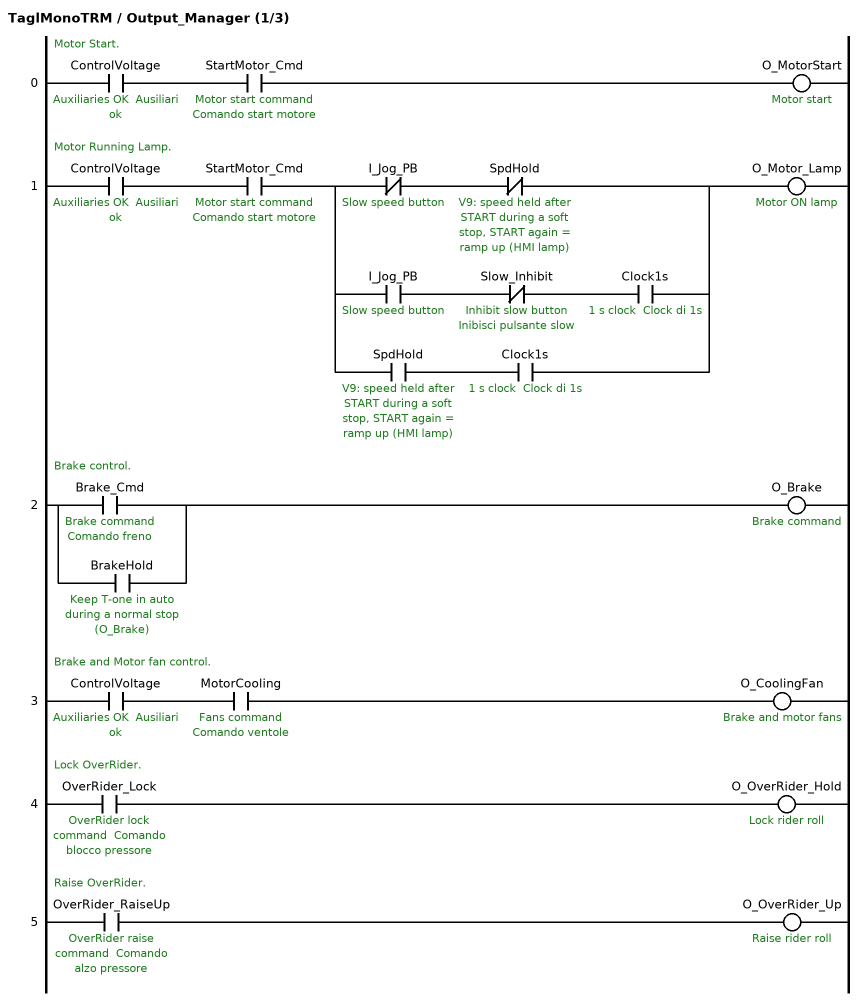
(* [picture p24: TaglMonoTRM / Output_Manager, rungs 0-5] *)
(* Rung 0: Motor Start. *)
O_MotorStart := ControlVoltage AND StartMotor_Cmd;
(* Rung 1: Motor Running Lamp. *)
O_Motor_Lamp := ControlVoltage AND StartMotor_Cmd AND ((NOT I_Jog_PB AND NOT SpdHold) OR (I_Jog_PB AND NOT Slow_Inhibit AND Clock1s) OR (SpdHold AND Clock1s));
(* Rung 2: Brake control. *)
O_Brake := Brake_Cmd OR BrakeHold;
(* Rung 3: Brake and Motor fan control. *)
O_CoolingFan := ControlVoltage AND MotorCooling;
(* Rung 4: Lock OverRider. *)
O_OverRider_Hold := OverRider_Lock;
(* Rung 5: Raise OverRider. *)
O_OverRider_Up := OverRider_RaiseUp;

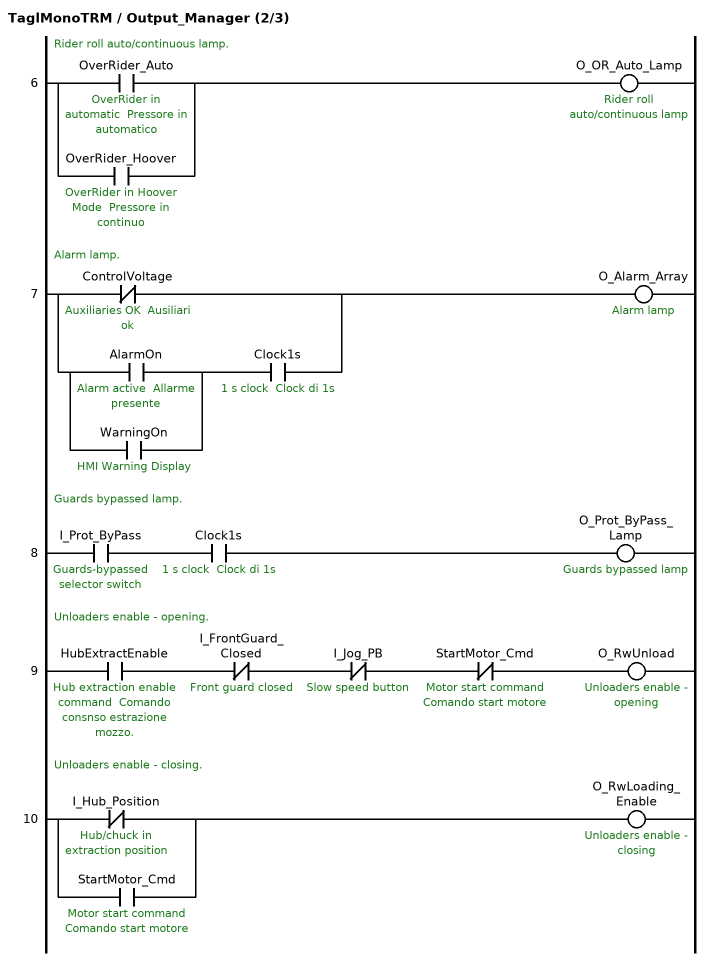
(* Rung 6: Rider roll auto/continuous lamp. *)
O_OR_Auto_Lamp := OverRider_Auto OR OverRider_Hoover;
(* Rung 7: Alarm lamp. *)
O_Alarm_Array := NOT ControlVoltage OR ((AlarmOn OR WarningOn) AND Clock1s);
(* Rung 8: Guards bypassed lamp. *)
O_Prot_ByPass_Lamp := I_Prot_ByPass AND Clock1s;
(* Rung 9: Unloaders enable - opening. *)
O_RwUnload := HubExtractEnable AND NOT I_FrontGuard_Closed AND NOT I_Jog_PB AND NOT StartMotor_Cmd;
(* Rung 10: Unloaders enable - closing. *)
O_RwLoading_Enable := NOT I_Hub_Position OR StartMotor_Cmd;

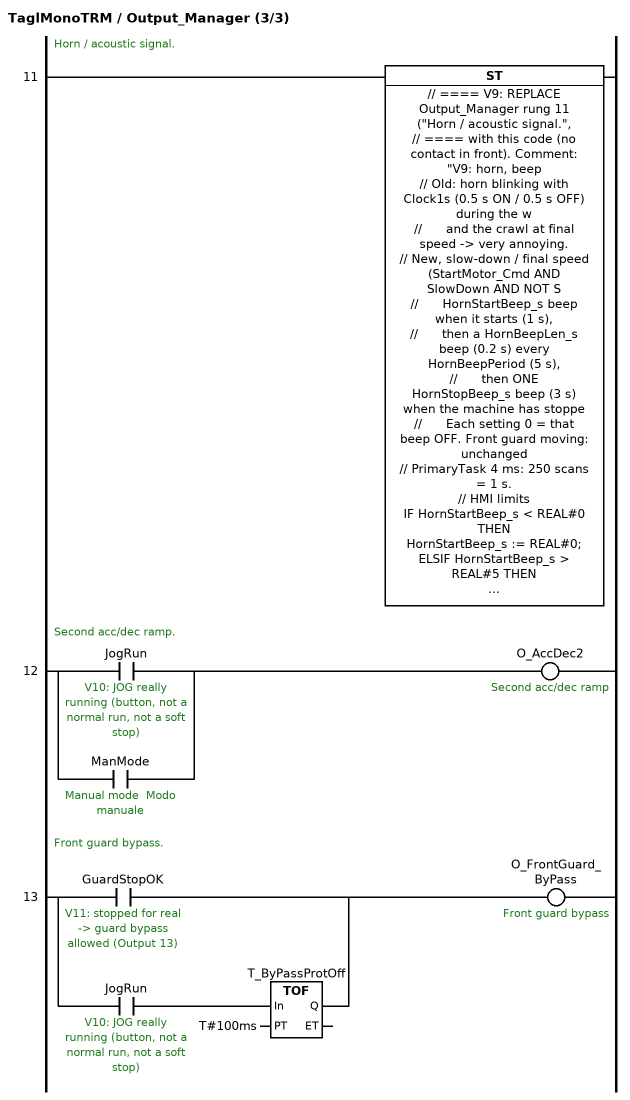
(* Rung 11: Horn / acoustic signal. *)
// ==== V9: REPLACE Output_Manager rung 11 ("Horn / acoustic signal.", ladder) by ONE ST rung
// ==== with this code (no contact in front). Comment: "V9: horn, beeps set on the HMI".
// Old: horn blinking with Clock1s (0.5 s ON / 0.5 s OFF) during the whole slow-down
//      and the crawl at final speed -> very annoying.
// New, slow-down / final speed (StartMotor_Cmd AND SlowDown AND NOT Stop):
//      HornStartBeep_s beep when it starts (1 s),
//      then a HornBeepLen_s beep (0.2 s) every HornBeepPeriod (5 s),
//      then ONE HornStopBeep_s beep (3 s) when the machine has stopped (< 2 m/min).
//      Each setting 0 = that beep OFF. Front guard moving: unchanged (Clock1s blinking).
// PrimaryTask 4 ms: 250 scans = 1 s.

// HMI limits

IF HornStartBeep_s < REAL#0 THEN
    HornStartBeep_s := REAL#0;
ELSIF HornStartBeep_s > REAL#5 THEN
    HornStartBeep_s := REAL#5;
END_IF;

IF HornBeepLen_s < REAL#0 THEN
    HornBeepLen_s := REAL#0;
ELSIF HornBeepLen_s > REAL#2 THEN
    HornBeepLen_s := REAL#2;
END_IF;

IF HornBeepPeriod < REAL#0 THEN
    HornBeepPeriod := REAL#0;
ELSIF (HornBeepPeriod > REAL#0) AND (HornBeepPeriod < HornBeepLen_s + REAL#0.5) THEN
    HornBeepPeriod := HornBeepLen_s + REAL#0.5;     // always a pause between beeps
ELSIF HornBeepPeriod > REAL#30 THEN
    HornBeepPeriod := REAL#30;
END_IF;

IF HornStopBeep_s < REAL#0 THEN
    HornStopBeep_s := REAL#0;
ELSIF HornStopBeep_s > REAL#10 THEN
    HornStopBeep_s := REAL#10;
END_IF;

HornStartScans := REAL_TO_INT(HornStartBeep_s * REAL#250);
HornLenScans   := REAL_TO_INT(HornBeepLen_s * REAL#250);
HornPer        := REAL_TO_INT(HornBeepPeriod * REAL#250);

// Slow-down / final speed beeps

HornRun := StartMotor_Cmd AND SlowDown AND NOT Stop;

IF HornRun THEN
    IF NOT HornRunMem THEN
        HornTicks := 0;                             // slow-down starts
    END_IF;
	
    IF HornTicks < 30000 THEN
        HornTicks := HornTicks + 1;
    END_IF;
	
    IF HornTicks <= HornStartScans THEN
        HornSlowBeep := TRUE;                       // start beep
        HornCnt := 0;
    ELSIF (HornPer > 0) AND (HornLenScans > 0) THEN
        HornCnt := HornCnt + 1;
        IF HornCnt >= HornPer THEN
            HornCnt := 0;
        END_IF;
		
        HornSlowBeep := (HornCnt >= HornPer - HornLenScans);   // beep at the end of each period
    ELSE
        HornSlowBeep := FALSE;                      // periodic beeps OFF
    END_IF;
ELSE
    HornTicks := 0;
    HornCnt := 0;
    HornSlowBeep := FALSE;
END_IF;

// End of a slow-down by a stop (auto stop, STOP button): one beep at standstill
// (Stop is set in Motor_Manager before StartMotor_Cmd drops on the next scan)

IF HornRunMem AND NOT HornRun AND (Stop OR NOT StartMotor_Cmd) THEN
    HornStopPend := TRUE;
END_IF;

IF StartMotor_Cmd AND NOT HornStartMem THEN
    HornStopPend := FALSE;                          // restarted: no stop beep
    HornStopTicks := 0;
END_IF;

HornStartMem := StartMotor_Cmd;

IF HornStopPend AND (Velocity_M_min < REAL#2) THEN
    HornStopPend := FALSE;
    HornStopTicks := REAL_TO_INT(HornStopBeep_s * REAL#250);
END_IF;

IF HornStopTicks > 0 THEN
    HornStopTicks := HornStopTicks - 1;
END_IF;

HornRunMem := HornRun;

// HMI test button: horn while pressed (machine stopped only)

O_AcousticSignal := (NOT I_FrontGuard_Closed AND NOT I_FrontGuard_Open AND Clock1s)
                    OR HornSlowBeep OR (HornStopTicks > 0)
                    OR (HornTest AND NOT StartMotor_Cmd);
(* Rung 12: Second acc/dec ramp. *)
O_AccDec2 := JogRun OR ManMode;
(* Rung 13: Front guard bypass. *)
T_ByPassProtOff(In := JogRun, PT := T#100ms);
O_FrontGuard_ByPass := GuardStopOK OR T_ByPassProtOff.Q;

(* Section AutoStop_Control: ladder, written here as Structured Text *)

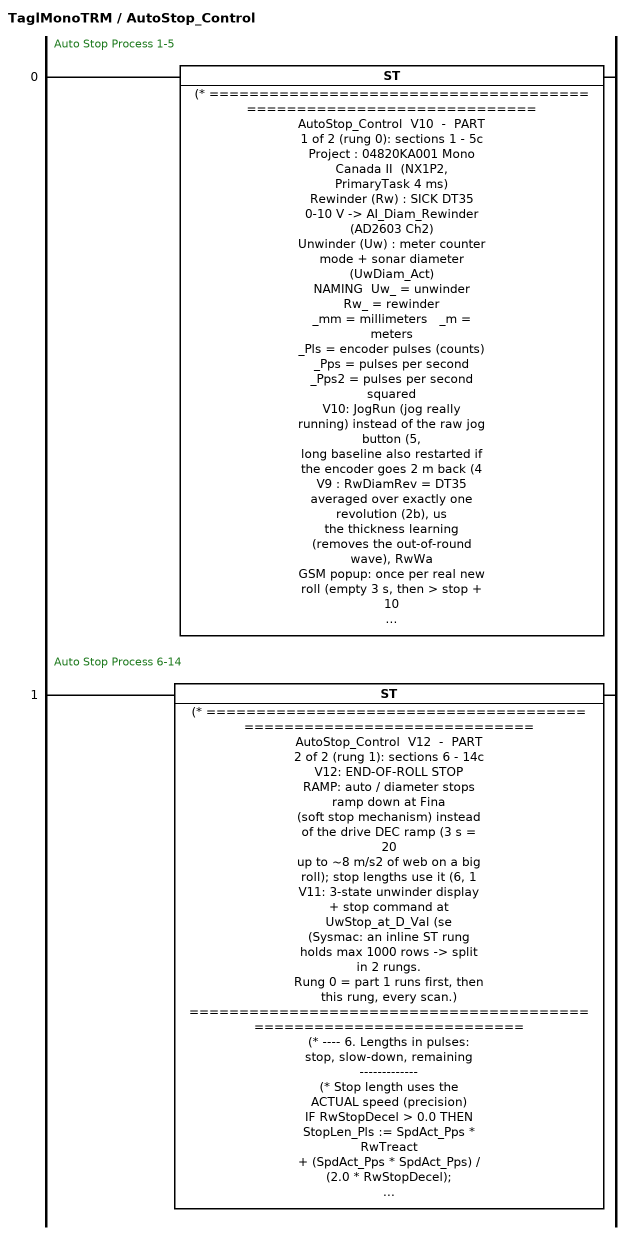
(* Rung 0: Auto Stop Process 1-5 *)
(* ==========================================================================
   AutoStop_Control  V10  -  PART 1 of 2 (rung 0): sections 1 - 5c
   Project : 04820KA001 Mono Canada II  (NX1P2, PrimaryTask 4 ms)
   Rewinder (Rw) : SICK DT35 0-10 V -> AI_Diam_Rewinder (AD2603 Ch2)
   Unwinder (Uw) : meter counter mode + sonar diameter (UwDiam_Act)

   NAMING  Uw_ = unwinder   Rw_ = rewinder
           _mm = millimeters   _m = meters
           _Pls = encoder pulses (counts)   _Pps = pulses per second
           _Pps2 = pulses per second squared

   V10: JogRun (jog really running) instead of the raw jog button (5, 5b);
          long baseline also restarted if the encoder goes 2 m back (4b).
   V9 : RwDiamRev = DT35 averaged over exactly one revolution (2b), used by
          the thickness learning (removes the out-of-round wave), RwWave_mm.
        GSM popup: once per real new roll (empty 3 s, then > stop + 100 mm
          for 3 s); NEW PAPER closes it (section 10).
        paper thickness: long-baseline learning (D^2 growth / length) from the
          start point, LOCKED at RwLockDiam (300 mm): no more change, no
          paper-change detection, until NEW PAPER / GSM popup YES (4b).
   V8 : = V7 + V7c unwinder DIAMETER slow-down follows the speed (6c),
          V7e ManMode slow-down model as before V7 (section 6),
          V7f S-curve extra length in the slow-down (section 6)
   V7 : FEED-FORWARD speed loop (Motor_Manager rung B): reference = set speed
        x RwRatioD / diameter along a ramp in real web mm/s2 (DecelWeb /
        AccelWeb), RwRatioD adapted slowly -> no hunting on big rolls.
        Section 6: slow-down length = one ramp at DecelWeb (FFEnable), else
        web coarse ramp + trim tail; learning only as fallback.
   v6y: rewinder AUTO stop (RwStopEnable) limits the work speed to
        RwAutoMaxSpd (500 m/min), taken over at standstill only; section 6
        uses the limited speed.
   v6x: new parent roll on the unwinder -> GsmAsk (HMI popup "did you change
        the paper?"); GsmAskYes forgets the learned thickness.
   v6w: paper thickness window is LENGTH-based instead of 10 s, modulated by
        the diameter (RwWinGrow_mm 2.5 mm of growth, 4 m .. RwWinLen_m 30 m):
        same accuracy at every speed and roll size; stopped window = dropped.
        ALARM RESET also clears LearnFailCnt / StopFailCnt (alarm 16).
   v6v: BrakeHold released on the SIGNED web speed (Velocity_M_min < 5),
        so a web pulled back after the stop releases the T-one at once.
   v6u: stop learning: a stop shorter than the reaction distance or faster
        than RwDecelMax_mm is ignored (not a fault). Only a too slow stop
        (< RwDecelMin_mm) counts toward alarm 16.
   v6t: rewinder slow-down fallback while the paper thickness is not
        learned: RwSlowReq at RwTargetDiam - RwSlowFallbackMm (30 mm).
   v6s: paper change: a learning window more than RwMatChangePct (25 %) away
        from RwMat_K is ignored once, taken directly the 2nd time in a row
        (automatic). RwMatReset (HMI "NEW PAPER") forgets RwMat_K.
   v6p: section 5c: RwLearnReset clears RwStopDecelK, RwStopDecel and
        RwSlowDecelK (the v6f seed that refilled RwStopDecelK is removed).
   v6l: previous value saved before every TEACH CORE (RwAxisDist_Prev,
          UwCoreDist_Prev, Retain) + UNDO buttons (RwTeachUndo,
          UwTeachUndo): swap current <-> previous. State 4 = RESTORED.
   v6k: unwinder TEACH CORE (Core_Measure) works like the rewinder one:
          same checks, 2 s stable with sonar AVERAGE, status UwTeachState.
          Replaces General rung 15 (one immediate sonar reading).
   v6j: TEACH CORE (section 14): HMI button RwTeachCore, empty core on the
          rewinder, machine stopped -> after 2 s stable:
          RwAxisDist := RwDist + RwCoreDiameter / 2. Status in RwTeachState.
   v6i: auto: pots scaled to WorkSpd_Max / FinalSpd_Max (Motor_Manager rung 6,
          Pot1_Mem / Pot2_Mem). ManMode keeps the raw pots (percent),
          so section 6 uses the raw pots in ManMode.
   v6h: BrakeHold keeps O_Brake (T-one "reel brake automatic") ON during a
          normal stop until the web is almost stopped (< 5 m/min, max 15 s).
          Before: T-one switched to "stop" with the run command, while the
          rewinder was decelerating hard -> unwinder overran, web on the
          floor (field 10/20/2026). Used in Output_Manager rung 2.
   v6g: slow-down AND stop decel proportional to the rewinder diameter.
          The ATV930 ramp is in Hz/s (motor = rewind shaft), so the web
          decel [mm/s2] = shaft decel x radius. Field data 10/20/2026:
          24 mm/s2 at 120 mm -> 90 mm/s2 at 600 mm.
          Learned: RwSlowDecelK, RwStopDecelK [mm/s2 per mm of diameter].
          Live:    RwSlowDecelLrn [mm/s2], RwStopDecel [pulses/s2] = K x DecelDiam.
   v6f: learn the REAL slow-down deceleration (section 5b) -> RwSlowDecelLrn
          (mm/s2). The ATV930 stretches its ramp with a heavy roll (no
          braking resistor), so the PLC ramp (DecelCoarse) was too
          optimistic: the stop came before final speed was reached.
          Priority in section 6: RwSlowDecel (manual) > RwSlowDecelLrn
          (learned) > DecelCoarse/DecelTrim model.
   v6e: GSM_Learned_OK (replaces global RwLearnFault): TRUE only when
          RwMat_K is learned, RwStopDecel is learned (if RwLearnStop) and
          there is no learning fault. Alarm 16 uses GSM_LearnFault.
   v6d: exact 100 ms tick (25 x 4 ms scan counter, the self-resetting
          TON ran ~104-108 ms -> speed ~4-8 % too high)
        standstill = <= 2 counts / 100 ms (encoder jitter)
        stop learning skipped after jog / manual / slow-button runs and
          when the auxiliaries drop (E-stop): RunWasJog, StopLearnValid
        work / final speed from the potentiometers in BOTH modes
          (Speed_Display / LowSpd_Display are not m/min in ManMode)
        slow-down length includes the DecelTrim tail inside the
          SpdDelta_Percent band (Motor_Manager rungs 14/15)
   v6c: learning supervision -> RwLearnFault (alarm 16), learned paper
          thickness RwThick_mm, plausibility limits for K and stop decel
   v6b: RwMaxSlowAtDiam display + RwMaxSlowFallback (slow-down warning
          while RwMat_K is not learned yet)
   v6 : consistent internal names, units in names.
        Globals renamed: RwRemain_m, RwStopLen_m, RwSlowLen_m,
                         RwSlowMargin_m, UwSlowMargin_m
   v5 : max diameter protection (always active), sensor plausibility,
        12SA5 master (section 9), alarms in section Alarms (ladder)
   v4b: AUTO interlock + single HMI display (SlowAtDisp / SlowAtMode)
   ========================================================================== *)

(* ---- 1. 100 ms tick, mm per encoder pulse ------------------------------ *)
(* v6d: 25 scans x 4 ms PrimaryTask = exactly 100 ms.                       *)
(*      Change 25 if the PrimaryTask period is changed.                    *)

TickCnt := TickCnt + 1;

IF TickCnt >= 25 THEN
    TickCnt := 0;
    Tick := TRUE;
ELSE
    Tick := FALSE;
END_IF;

IF (Encoder_Pulse > 0) AND (EncoderWheel_Circumf > 0.0) THEN
    MmPerPulse := EncoderWheel_Circumf / (INT_TO_REAL(Encoder_Pulse) * 4.0);
ELSE
    MmPerPulse := 0.0;
END_IF;

(* ---- 2. Rewinder DT35 -> filtered distance -> diameter ----------------- *)

RwDistRaw_mm := RwDist0V + (INT_TO_REAL(AI_Diam_Rewinder) / 4000.0)
                * (RwDist10V - RwDist0V);

IF Tick THEN
    IF NOT RwFiltInit THEN
        RwDist := RwDistRaw_mm;
        RwFiltInit := TRUE;
    ELSE
        RwDist := RwDist + RwFilter_K * (RwDistRaw_mm - RwDist);
    END_IF;
END_IF;

RwSensFault := (AI_Diam_Rewinder < RwRawMin) OR (AI_Diam_Rewinder > RwRawMax)
               OR (RwDist > RwAxisDist);

RwDiam := 2.0 * (RwAxisDist - RwDist);

IF RwDiam < 0.0 THEN
    RwDiam := 0.0;
END_IF;

(* ---- 2b. V9: diameter averaged over exactly ONE revolution -------------- *)
(* The out-of-round roll gives a wave at the rotation frequency (seen in   *)
(* the 10/29 traces: 2.4 Hz at 444 m/min / 973 mm). Averaging the raw     *)
(* DT35 distance over exactly one revolution cancels it (and all its      *)
(* harmonics), whatever the phase -> no shaft position sensor needed:     *)
(* one revolution = PI x D of web on the encoder. Each scan is weighted   *)
(* by its encoder pulses = by roll ANGLE, so ramps and standstill do not  *)
(* bias it (stopped: nothing added). Used only by the thickness learning. *)
(* RwWave_mm = peak-peak diameter wave in the last revolution (HMI).      *)

RevDP := ABS(Encoder_Pos - RevPrevPos);
RevPrevPos := Encoder_Pos;

IF RwSensFault OR (MmPerPulse <= 0.0) OR (RwDiam < 50.0) OR (RevDP > 100000) THEN
    RevW := 0.0;
    RevSum := 0.0;
    RwDiamRevOk := RwDiamRevOk AND NOT RwSensFault;
ELSIF RevDP > 0 THEN
	
    IF RevW <= 0.0 THEN
        RevMin := RwDistRaw_mm;
        RevMax := RwDistRaw_mm;
    END_IF;
	
    RevSum := RevSum + RwDistRaw_mm * DINT_TO_REAL(RevDP);
    RevW := RevW + DINT_TO_REAL(RevDP);
	
    IF RwDistRaw_mm < RevMin THEN
        RevMin := RwDistRaw_mm;
    END_IF;
	
    IF RwDistRaw_mm > RevMax THEN
        RevMax := RwDistRaw_mm;
    END_IF;
	
    IF RevW >= 3.14159 * RwDiam / MmPerPulse THEN
        RwDiamRev := 2.0 * (RwAxisDist - RevSum / RevW);
        RwWave_mm := 2.0 * (RevMax - RevMin);
        RwDiamRevOk := TRUE;
        RevW := 0.0;
        RevSum := 0.0;
    END_IF;
END_IF;

(* v6g: diameter used by the decel model (last valid on sensor fault)      *)

IF NOT RwSensFault THEN
    DecelDiam := RwDiam;
ELSE
    DecelDiam := RwLastValidDiam;
END_IF;

IF DecelDiam < 100.0 THEN
    DecelDiam := 100.0;                             (* core *)
END_IF;

(* ---- 3. Actual speed from encoder, 100 ms window ----------------------- *)

IF Tick THEN
	
    IF NOT SpdInit THEN
        EncPrev := Encoder_Pos;
        SpdInit := TRUE;
    END_IF;
	
    SpdAct_Pps := DINT_TO_REAL(ABS(Encoder_Pos - EncPrev)) * 10.0;
    EncPrev := Encoder_Pos;
END_IF;

RwSpeed := SpdAct_Pps * MmPerPulse * 0.06;          (* m/min *)

(* ---- 4a. v6s: NEW PAPER button: forget the learned thickness ----------- *)
(* RwMat_K = 0 -> the first valid 10 s window sets it directly.            *)
(* HMI momentary button: must be HELD 3 s, then the reset is done once and *)
(* the PLC clears the bit (HMI lamp goes off = done).                      *)

T_MatReset(In := RwMatReset, PT := T#3s);

IF T_MatReset.Q THEN
    RwMat_K := 0.0;
    LearnFailCnt := 0;
    MatChangeCnt := 0;
    RwMatLocked := FALSE;                           (* V9 *)
    LongActive := FALSE;
    GsmAsk := FALSE;                                (* V9: NEW PAPER answers the popup *)
    GsmArmed := FALSE;
    RwMatReset := FALSE;
END_IF;

(* ---- 4b. V9: long-baseline thickness learning + LOCK ------------------- *)
(* From the start point (first run after NEW PAPER / GSM YES / power-on    *)
(* while not locked): K = (D^2 - D0^2) / (2 x pulses). The waving of the   *)
(* roll (+/-0.4 mm) only matters at the two ends, so the error falls with  *)
(* the growth (50 mm growth: ~1 %). After 20 mm growth it replaces the     *)
(* 30 m windows. At RwLockDiam (and >= RwLockMinGrow_mm growth) the value *)
(* is LOCKED (Retain): windows and paper-change detection stop.            *)
(* RwLockDiam = 0 -> never locked (windows + long baseline as learning).   *)

IF Tick AND NOT RwMatLocked THEN
	
    IF LongActive AND (RwDiamRev < LongStartD - 30.0) AND RwDiamRevOk THEN
        LongActive := FALSE;                        (* new core: restart *)
    END_IF;
	
    IF Encoder_Reset OR (Encoder_Pos < LongStartPos - 20000) THEN
        LongActive := FALSE;                        (* metre counter reset / 2 m back *)
    END_IF;
	
    IF NOT LongActive AND O_MotorStart AND RwDiamRevOk
       AND (RwDiamRev > 0.0) THEN
        LongStartPos := Encoder_Pos;
        LongStartD := RwDiamRev;
        LongActive := TRUE;
    END_IF;
	
    LongValid := FALSE;
	
    IF LongActive AND RwDiamRevOk AND (MmPerPulse > 0.0) THEN
        LongGrow_mm := RwDiamRev - LongStartD;
        LongPls := DINT_TO_REAL(ABS(Encoder_Pos - LongStartPos));
		
        IF (LongGrow_mm >= 20.0) AND (LongPls > 0.0) THEN
            LongK := (RwDiamRev * RwDiamRev - LongStartD * LongStartD) / (2.0 * LongPls);
            LongThick_mm := LongK * 3.14159 / (2.0 * MmPerPulse);
			
            IF (LongThick_mm >= RwThickMin_mm) AND (LongThick_mm <= RwThickMax_mm) THEN
                LongValid := TRUE;
                RwMat_K := LongK;
                MatChangeCnt := 0;
                LearnFailCnt := 0;
				
                IF (RwLockDiam > 0.0) AND (RwDiamRev >= RwLockDiam)
                   AND (LongGrow_mm >= RwLockMinGrow_mm) THEN
                    RwMatLocked := TRUE;            (* solid from now on *)
                    LongActive := FALSE;
                END_IF;
            END_IF;
        END_IF;
    END_IF;
END_IF;

IF RwMatLocked THEN
    LongValid := FALSE;
    LearnFailCnt := 0;                              (* no thickness alarm *)
END_IF;

(* ---- 4. Learn material factor  K = dDiam/dPulse * Diam ----------------- *)

IF Tick THEN
    LearnWinTicks := LearnWinTicks + 1;
	
    IF NOT LearnInit THEN
        LearnWinStartPos := Encoder_Pos;  LearnWinStartDiam := RwDiamRev;  (* V9 *)
        LearnWinTicks := 0;
        LearnWinRunning := O_MotorStart;
        LearnInit := TRUE;
    ELSE
        LearnWinRunning := LearnWinRunning AND O_MotorStart;
        (* v6w: LENGTH-based window, modulated by the diameter: closes    *)
        (* when the roll should have grown RwWinGrow_mm (2.5 mm), so the  *)
        (* accuracy vs DT35 noise is the same at every speed and size.    *)
        (* Pulses = growth x diameter / K (K = learned RwMat_K).          *)
        (* Limits: min 4 m, max RwWinLen_m (30 m). K not learned: max.    *)
        (* Motor stopped during the window -> window dropped (no fault).  *)
		
        IF MmPerPulse > 0.0 THEN
            IF (RwMat_K > 0.0) AND (RwWinGrow_mm > 0.0) THEN
                LearnWinLen_Pls := RwWinGrow_mm * MAX(RwDiam, REAL#100.0) / RwMat_K;
            ELSE
                LearnWinLen_Pls := RwWinLen_m * 1000.0 / MmPerPulse;
            END_IF;
			
            IF LearnWinLen_Pls < 4000.0 / MmPerPulse THEN
                LearnWinLen_Pls := 4000.0 / MmPerPulse;              (* 4 m *)
            END_IF;
			
            IF (RwWinLen_m > 0.0)
               AND (LearnWinLen_Pls > RwWinLen_m * 1000.0 / MmPerPulse) THEN
                LearnWinLen_Pls := RwWinLen_m * 1000.0 / MmPerPulse;
            END_IF;
        ELSE
            LearnWinLen_Pls := 300000.0;
        END_IF;
		
        IF (DINT_TO_REAL(ABS(Encoder_Pos - LearnWinStartPos)) >= LearnWinLen_Pls)
           OR NOT LearnWinRunning THEN
            LearnWin_Pls := ABS(Encoder_Pos - LearnWinStartPos);
            LearnWinDiamDelta := RwDiamRev - LearnWinStartDiam;  (* V9 *)
            (* A window SHOULD learn: ran all the time, enough length,  *)
            (* DT35 OK. Then it must give a plausible paper thickness. *)
			
            IF LearnWinRunning AND (LearnWin_Pls >= RwMinPulses)
               AND NOT RwSensFault
               AND NOT RwMatLocked AND NOT LongValid      (* V9 *)
               AND RwDiamRevOk AND (LearnWinStartDiam > 0.0) THEN
                LearnWinOk := FALSE;
				
                IF (LearnWinDiamDelta > 0.0) AND (MmPerPulse > 0.0) THEN
                    MatK_Window := (LearnWinDiamDelta / DINT_TO_REAL(LearnWin_Pls))
                                   * ((RwDiamRev + LearnWinStartDiam) / 2.0);
                    (* K = 2 * thickness * mm-per-pulse / PI          *)
                    ThickWin_mm := MatK_Window * 3.14159 / (2.0 * MmPerPulse);
					
                    IF (ThickWin_mm >= RwThickMin_mm)
                       AND (ThickWin_mm <= RwThickMax_mm) THEN
                        LearnWinOk := TRUE;
						
                        IF RwMat_K <= 0.0 THEN
                            RwMat_K := MatK_Window;
                            MatChangeCnt := 0;
                        ELSIF (RwMatChangePct > 0.0)
                              AND (ABS(MatK_Window - RwMat_K)
                                   > RwMat_K * RwMatChangePct / 100.0) THEN
                            (* v6s: far from the learned value: 1 window = ignored *)
                            (* (outlier), 2 in a row = paper changed -> take it.  *)
                            MatChangeCnt := MatChangeCnt + 1;
							
                            IF MatChangeCnt >= 2 THEN
                                RwMat_K := MatK_Window;
                                MatChangeCnt := 0;
                            END_IF;
                        ELSE
                            MatChangeCnt := 0;
                            RwMat_K := RwMat_K + RwLearn_K * (MatK_Window - RwMat_K);
                        END_IF;
                    END_IF;
                END_IF;
				
                IF LearnWinOk THEN
                    LearnFailCnt := 0;
                ELSIF LearnFailCnt < 1000 THEN
                    LearnFailCnt := LearnFailCnt + 1;  (* no growth / implausible *)
                END_IF;
            END_IF;
            LearnWinStartPos := Encoder_Pos;  LearnWinStartDiam := RwDiamRev;  (* V9 *)
            LearnWinTicks := 0;
            LearnWinRunning := O_MotorStart;
        END_IF;
    END_IF;
END_IF;

(* ---- 5. Learn real stop deceleration on every stop --------------------- *)
(* v6d: a run with jog / manual / slow button uses the 2nd ramp (O_AccDec2) *)
(*      -> its stop must not be learned. Latched for the whole run because  *)
(*      the jog button is already released on the stop edge.                  *)

IF O_MotorStart AND NOT MotorRunMem THEN            (* start edge *)
    RunWasJog := FALSE;
END_IF;

IF O_MotorStart AND (ManMode OR JogRun) THEN
    RunWasJog := TRUE;
END_IF;

IF MotorRunMem AND NOT O_MotorStart THEN            (* stop command edge *)
    StopMeasActive := TRUE;
    StopStartPos := Encoder_Pos;
    StopStartSpd_Pps := SpdAct_Pps;
    StopStartDiam := DecelDiam;
    StandstillTicks := 0;
    (* STOP button and automatic stop take the same path (drive DI1 and    *)
    (* O_Brake -> T-one drop together, electrical plan sheets 1/9/15),     *)
    (* so both are learned.                                                *)
    StopLearnValid := ControlVoltage AND NOT RunWasJog AND NOT ManMode;
END_IF;

MotorRunMem := O_MotorStart;

IF O_MotorStart THEN
    StopMeasActive := FALSE;                        (* restarted: abort *)
ELSIF StopMeasActive AND Tick THEN
	
    IF NOT ControlVoltage THEN
        StopLearnValid := FALSE;                    (* E-stop during the stop *)
    END_IF;
	
    IF SpdAct_Pps <= 20.0 THEN                      (* <= 2 counts / 100 ms *)
        StandstillTicks := StandstillTicks + 1;
    ELSE
        StandstillTicks := 0;
    END_IF;
	
    IF StandstillTicks >= 3 THEN                    (* standstill 300 ms *)
        StopMeasActive := FALSE;
        StopMeas_Pls := DINT_TO_REAL(ABS(Encoder_Pos - StopStartPos));
		
        IF RwLearnStop AND StopLearnValid
           AND (StopStartSpd_Pps * MmPerPulse * 0.06 >= RwMinLearnSpd) THEN
            (* This stop SHOULD learn: result must be plausible       *)
            (* v6u: a stop shorter than the reaction distance, or     *)
            (* faster than RwDecelMax_mm, is NOT a fault: the web      *)
            (* stopped within a few mm, nothing to learn (trace        *)
            (* 10/28/2026: 23 m/min -> stopped in 102 pulses = 10 mm). *)
            (* Only a too SLOW stop (< RwDecelMin_mm) counts as fail.  *)
            StopLearnOk := FALSE;
			
            IF StopMeas_Pls > StopStartSpd_Pps * RwTreact THEN
                StopDecelMeas := (StopStartSpd_Pps * StopStartSpd_Pps)
                                 / (2.0 * (StopMeas_Pls - StopStartSpd_Pps * RwTreact));
                StopDecelMeas_mm := StopDecelMeas * MmPerPulse;  (* mm/s2 *)
				
                IF (StopDecelMeas_mm >= RwDecelMin_mm)
                   AND (StopDecelMeas_mm <= RwDecelMax_mm) THEN
                    StopLearnOk := TRUE;
                    (* v6g: learn per mm of diameter *)
                    DecelK_Meas := StopDecelMeas_mm / ((StopStartDiam + DecelDiam) / 2.0);
					
                    IF RwStopDecelK <= 0.0 THEN
                        RwStopDecelK := DecelK_Meas;
                    ELSE
                        RwStopDecelK := RwStopDecelK + 0.3 * (DecelK_Meas - RwStopDecelK);
                    END_IF;
					
                    StopFailCnt := 0;
                ELSIF StopDecelMeas_mm < RwDecelMin_mm THEN
					
                    IF StopFailCnt < 1000 THEN
                        StopFailCnt := StopFailCnt + 1;    (* stop too long *)
                    END_IF;
                END_IF;                                    (* too fast: ignored *)
            END_IF;                                        (* too short: ignored *)
        END_IF;
    END_IF;
END_IF;

(* ---- 5b. v6f: learn real slow-down deceleration ----------------------- *)
(* From the SlowDown edge (at speed) until final speed is reached, or     *)
(* until the stop comes first. a = (v0^2 - v1^2) / (2 * distance).         *)
(* Not learned in jog / manual / slow button (2nd ramp).                   *)

IF SlowDown AND NOT SlowMem AND O_MotorStart
   AND NOT ManMode AND NOT JogRun
   AND (SpdAct_Pps > SpdFinal_Pps + SpdBand_Pps) THEN
    SlowMeasActive := TRUE;
    SlowStartPos := Encoder_Pos;
    SlowStartSpd_Pps := SpdAct_Pps;
    SlowStartDiam := DecelDiam;
END_IF;
SlowMem := SlowDown;

IF SlowMeasActive THEN
	
    IF NOT SlowDown OR ManMode OR JogRun THEN
        SlowMeasActive := FALSE;                    (* aborted *)
    ELSIF Tick AND ((SpdAct_Pps <= SpdFinal_Pps + 0.25 * SpdBand_Pps)
                    OR NOT O_MotorStart) THEN       (* final reached or stopped *)
        SlowMeasActive := FALSE;
        SlowMeas_Pls := DINT_TO_REAL(ABS(Encoder_Pos - SlowStartPos));
		
        IF (SlowMeas_Pls > 0.0) AND (MmPerPulse > 0.0)
           AND ((SlowStartSpd_Pps - SpdAct_Pps) * MmPerPulse * 0.06 >= 10.0) THEN
            SlowDecelMeas_mm := (SlowStartSpd_Pps * SlowStartSpd_Pps
                                 - SpdAct_Pps * SpdAct_Pps)
                                / (2.0 * SlowMeas_Pls) * MmPerPulse;  (* mm/s2 *)
								
            IF (SlowDecelMeas_mm >= RwDecelMin_mm)
               AND (SlowDecelMeas_mm <= RwDecelMax_mm) THEN
                (* v6g: learn per mm of diameter *)
                DecelK_Meas := SlowDecelMeas_mm / ((SlowStartDiam + DecelDiam) / 2.0);
				
                IF RwSlowDecelK <= 0.0 THEN
                    RwSlowDecelK := DecelK_Meas;
                ELSE
                    RwSlowDecelK := RwSlowDecelK + 0.5 * (DecelK_Meas - RwSlowDecelK);
                END_IF;
            END_IF;
        END_IF;
    END_IF;
END_IF;

(* ---- 5c. v6g: live decels = learned K x current diameter -------------- *)
(* v6p: the one-time v6f seed is removed (it re-filled RwStopDecelK from    *)
(* RwStopDecel, so the learning could never be reset).                     *)
(* RwLearnReset (HMI / Watch tab, PLC resets it): clear the learned decels. *)
(* Both are re-learned at the next auto slow-down / stop >= RwMinLearnSpd.  *)

IF RwLearnReset THEN
    RwStopDecelK := 0.0;
    RwStopDecel := 0.0;
    RwSlowDecelK := 0.0;
    StopFailCnt := 0;
    RwLearnReset := FALSE;
END_IF;

IF (RwStopDecelK > 0.0) AND (MmPerPulse > 0.0) THEN
    RwStopDecel := RwStopDecelK * DecelDiam / MmPerPulse;      (* pulses/s2 *)
END_IF;

IF RwSlowDecelK > 0.0 THEN
    RwSlowDecelLrn := RwSlowDecelK * DecelDiam;                (* mm/s2 *)
ELSE
    RwSlowDecelLrn := 0.0;
END_IF;
(* Rung 1: Auto Stop Process 6-14 *)
(* ==========================================================================
   AutoStop_Control  V12  -  PART 2 of 2 (rung 1): sections 6 - 14c
   V12: END-OF-ROLL STOP RAMP: auto / diameter stops ramp down at FinalStopDecel
        (soft stop mechanism) instead of the drive DEC ramp (3 s = 20 Hz/s,
        up to ~8 m/s2 of web on a big roll); stop lengths use it (6, 11b).
   V11: 3-state unwinder display + stop command at UwStop_at_D_Val (section 8).
   (Sysmac: an inline ST rung holds max 1000 rows -> split in 2 rungs.
    Rung 0 = part 1 runs first, then this rung, every scan.)
   ========================================================================== *)

(* ---- 6. Lengths in pulses: stop, slow-down, remaining ------------------ *)
(* Stop length uses the ACTUAL speed (precision)                           *)

IF RwStopDecel > 0.0 THEN
    StopLen_Pls := SpdAct_Pps * RwTreact
                   + (SpdAct_Pps * SpdAct_Pps) / (2.0 * RwStopDecel);
ELSE
    StopLen_Pls := SpdAct_Pps * (RwTreact + RwTstopDef / 2.0);
END_IF;

(* V12: end-of-roll stop ramp at FinalStopDecel (web mm/s2) + S-curve    *)

IF (FinalStopDecel > 0.0) AND FFEnable AND NOT ManMode AND (MmPerPulse > 0.0) THEN
    StopLen_Pls := SpdAct_Pps * RwTreact
                   + (SpdAct_Pps * SpdAct_Pps) / (2.0 * FinalStopDecel / MmPerPulse)
                   + SpdAct_Pps * 0.5 * SCurveTime;
END_IF;

StopLen_Pls := StopLen_Pls * RwTrim;

(* Slow-down uses SpdRef = MAX(actual, work-speed setpoint):               *)
(* stable value, shown to the operator even before start                   *)

SlowLenBase_Pls := 0.0;  RwSlowLen_Pls := 0.0;  UwSlowLen_Pls := 0.0;

IF MmPerPulse > 0.0 THEN
    (* v6f: manual > learned > PLC ramp model                           *)
    (* V7: manual > feed-forward (one ramp at DecelWeb, real web mm/s2)  *)
    (*     > old loop with web ramps (coarse DecelWeb + trim tail)       *)
    (*     > learned > old PLC ramp model                                *)
	
    IF RwSlowDecel > 0.0 THEN
        SlowDecel_Pps2 := RwSlowDecel / MmPerPulse;
        SlowOneRamp := TRUE;
    ELSIF FFEnable AND (DecelWeb > 0.0) AND (WebRatio > 0.0) AND NOT ManMode THEN
        SlowDecel_Pps2 := DecelWeb / MmPerPulse;
        SlowOneRamp := TRUE;
    ELSIF (DecelWeb > 0.0) AND (WebRatio > 0.0) AND NOT ManMode THEN  (* V7e *)
        SlowDecel_Pps2 := DecelWeb / MmPerPulse;
        SlowOneRamp := FALSE;
    ELSIF RwSlowDecelLrn > 0.0 THEN
        SlowDecel_Pps2 := RwSlowDecelLrn / MmPerPulse;  (* real, incl. trim tail *)
        SlowOneRamp := TRUE;
    ELSE
        SlowDecel_Pps2 := DecelCoarse * 250.0 / MmPerPulse; (* 1 = 250 mm/s2 *)
        SlowOneRamp := FALSE;
    END_IF;
	
    (* v6d: DecelTrim ramp used inside the +/- SpdDelta_Percent band *)
	
    IF (DecelTrim > 0.0) AND (WebRatio > 0.0) AND (Vel_Max_mms > 0.0) THEN
        (* V7: trim ramp (reference units) converted to the real web decel *)
        TrimDecel_Pps2 := DecelTrim * 1000000.0 / (0.06 * WebRatio * Vel_Max_mms)
                          / MmPerPulse;
    ELSIF DecelTrim > 0.0 THEN
        TrimDecel_Pps2 := DecelTrim * 250.0 / MmPerPulse;
    ELSE
        TrimDecel_Pps2 := SlowDecel_Pps2;
    END_IF;
	
    SpdBand_Pps := SpdDelta_Percent * 1000.0 / 60.0 / MmPerPulse;

    (* v6d: speeds from the potentiometers, valid in auto AND ManMode     *)
    (*      (m/min = Pot / Input_Ratio, same as Motor_Manager rung 8)     *)
	
    IF (Input_Ratio > 0.0) AND ManMode THEN
        (* v6i: ManMode drives the inverter with the raw pots (rung 17) *)
        SpdFinal_Pps := INT_TO_REAL(Pot2_Slow_Velocity) / Input_Ratio * 1000.0 / 60.0 / MmPerPulse;
        SpdWork_Pps  := INT_TO_REAL(Pot1_Work_Velocity) / Input_Ratio * 1000.0 / 60.0 / MmPerPulse;
    ELSIF Input_Ratio > 0.0 THEN
        SpdFinal_Pps := INT_TO_REAL(Pot2_Mem) / Input_Ratio * 1000.0 / 60.0 / MmPerPulse;
        SpdWork_Pps  := INT_TO_REAL(Pot1_Mem) / Input_Ratio * 1000.0 / 60.0 / MmPerPulse;
    ELSE
        SpdFinal_Pps := LowSpd_Display * 1000.0 / 60.0 / MmPerPulse;
        SpdWork_Pps  := Speed_Display  * 1000.0 / 60.0 / MmPerPulse;
    END_IF;
	
    (* v6y: rewinder AUTO stop -> work speed limited to RwAutoMaxSpdAct *)
    (* (limit + value taken over only at standstill, Motor_Manager rung 5) *)
	
    IF RwAutoLimAct AND NOT ManMode
       AND (SpdWork_Pps > RwAutoMaxSpdAct * 1000.0 / 60.0 / MmPerPulse) THEN
        SpdWork_Pps := RwAutoMaxSpdAct * 1000.0 / 60.0 / MmPerPulse;
    END_IF;
	
    SpdRef_Pps := MAX(SpdAct_Pps, SpdWork_Pps);

    IF RwStopDecel > 0.0 THEN
        StopLenFinal_Pls := SpdFinal_Pps * RwTreact
                            + (SpdFinal_Pps * SpdFinal_Pps) / (2.0 * RwStopDecel);
    ELSE
        StopLenFinal_Pls := SpdFinal_Pps * (RwTreact + RwTstopDef / 2.0);
    END_IF;

    (* V12: final stop from the final speed on the end-of-roll ramp *)
	
    IF (FinalStopDecel > 0.0) AND FFEnable AND NOT ManMode THEN
        StopLenFinal_Pls := SpdFinal_Pps * RwTreact
                            + (SpdFinal_Pps * SpdFinal_Pps) / (2.0 * FinalStopDecel / MmPerPulse)
                            + SpdFinal_Pps * 0.5 * SCurveTime;
    END_IF;

    SlowLenBase_Pls := StopLenFinal_Pls * RwTrim;
	
    IF (SpdRef_Pps > SpdFinal_Pps) AND (SlowDecel_Pps2 > 0.0) THEN
		
        IF SlowOneRamp OR (TrimDecel_Pps2 <= 0.0) THEN
            (* manual or learned decel: one constant ramp *)
            SlowLenBase_Pls := SlowLenBase_Pls
                + (SpdRef_Pps * SpdRef_Pps - SpdFinal_Pps * SpdFinal_Pps)
                  / (2.0 * SlowDecel_Pps2);
        ELSE
            (* auto: coarse ramp down to the band, trim ramp inside it *)
            SpdKnee_Pps := SpdFinal_Pps + SpdBand_Pps;
			
            IF SpdRef_Pps > SpdKnee_Pps THEN
                SlowLenBase_Pls := SlowLenBase_Pls
                    + (SpdRef_Pps * SpdRef_Pps - SpdKnee_Pps * SpdKnee_Pps)
                      / (2.0 * SlowDecel_Pps2)
                    + (SpdKnee_Pps * SpdKnee_Pps - SpdFinal_Pps * SpdFinal_Pps)
                      / (2.0 * TrimDecel_Pps2);
            ELSE
                SlowLenBase_Pls := SlowLenBase_Pls
                    + (SpdRef_Pps * SpdRef_Pps - SpdFinal_Pps * SpdFinal_Pps)
                      / (2.0 * TrimDecel_Pps2);
            END_IF;
        END_IF;
    END_IF;

    (* V7f: S-curve rounding: the slow-down ends SCurveTime later ->      *)
    (*      extra length = (SpdRef - SpdFinal) / 2 x SCurveTime            *)
	
    IF FFEnable AND NOT ManMode AND (RwSlowDecel <= 0.0) AND (DecelWeb > 0.0)
       AND (WebRatio > 0.0) AND (SCurveTime > 0.0)
       AND (SpdRef_Pps > SpdFinal_Pps) THEN
        SlowLenBase_Pls := SlowLenBase_Pls
                           + (SpdRef_Pps - SpdFinal_Pps) * 0.5 * SCurveTime;
    END_IF;

    RwSlowLen_Pls := SlowLenBase_Pls + RwSlowMargin_m * 1000.0 / MmPerPulse;

    IF UwSlowMargin_m > 0.0 THEN
        UwMarginUsed_m := UwSlowMargin_m;
    ELSE
        UwMarginUsed_m := RwSlowMargin_m;
    END_IF;
	
    UwSlowLen_Pls := SlowLenBase_Pls + UwMarginUsed_m * 1000.0 / MmPerPulse;
END_IF;

IF RwDiam >= RwTargetDiam THEN
    RwRemain_Pls := 0.0;
ELSIF RwMat_K > 0.0 THEN
    RwRemain_Pls := (RwTargetDiam * RwTargetDiam - RwDiam * RwDiam)
                    / (2.0 * RwMat_K);
ELSE
    RwRemain_Pls := 1.0E9;                          (* K not learned: plain target *)
END_IF;

RwRemain_m  := RwRemain_Pls  * MmPerPulse / 1000.0;
RwStopLen_m := StopLen_Pls   * MmPerPulse / 1000.0;
RwSlowLen_m := RwSlowLen_Pls * MmPerPulse / 1000.0;

(* ---- 6b. Live operator displays ---------------------------------------- *)
(* Rewinder: diameter where slow-down / stop command will happen           *)

IF RwMat_K > 0.0 THEN
    SqrtArg := RwTargetDiam * RwTargetDiam - 2.0 * RwMat_K * RwSlowLen_Pls;
    IF SqrtArg > 0.0 THEN
        RwSlow_at_D_Val := SQRT(SqrtArg);
    ELSE
        RwSlow_at_D_Val := 0.0;
    END_IF;
	
    SqrtArg := RwTargetDiam * RwTargetDiam - 2.0 * RwMat_K * StopLen_Pls;
	
    IF SqrtArg > 0.0 THEN
        RwStop_at_D_Val := SQRT(SqrtArg);
    ELSE
        RwStop_at_D_Val := 0.0;
    END_IF;
ELSE
    (* v6t: thickness not learned: fixed slow-down point before the target *)
	
    IF RwUseSlow AND (RwSlowFallbackMm > 0.0) THEN
        RwSlow_at_D_Val := RwTargetDiam - RwSlowFallbackMm;
    ELSE
        RwSlow_at_D_Val := RwTargetDiam;
    END_IF;
    RwStop_at_D_Val := RwTargetDiam;
END_IF;

(* Unwinder: meter count where the slow-down will start                   *)

IF MmPerPulse > 0.0 THEN
    UwSlow_at_M_Val := UwStop_at_M_Val - UwSlowLen_Pls * MmPerPulse / 1000.0;
ELSE
    UwSlow_at_M_Val := UwStop_at_M_Val;
END_IF;

IF UwSlow_at_M_Val < 0.0 THEN
    UwSlow_at_M_Val := 0.0;
END_IF;

(* Unwinder slow-down request, latched                                     *)

IF (Current_Metre < UwSlow_at_M_Val - 50.0) OR (UwStop_at_M_Val <= 0.0) THEN
    UwSlow_at_M_Req := FALSE;                             (* counter reset / longer roll *)
END_IF;

IF (UwStop_at_M_Val > 0.0) AND (Current_Metre >= UwSlow_at_M_Val) THEN
    UwSlow_at_M_Req := TRUE;
END_IF;

(* ---- 6c. V7c: unwinder DIAMETER slow-down follows the speed ----------- *)
(* Works without AutoStop (only Measure_ON, like General rung 16).         *)
(* Paper left above the stop diameter, in pulses:                          *)
(*     (UwDiam_Act^2 - UwStopDiam_Limit^2) / (2 x RwMat_K)                        *)
(* (same paper as the rewinder -> same learned K). Slow down when it is    *)
(* shorter than UwSlowLen_Pls = decel from the speed (DecelWeb) + final    *)
(* stop + UwSlowMargin_m. Solved for the diameter:                         *)
(*     UwSlowDiamCalc = SQRT(UwStopDiam_Limit^2 + 2 x RwMat_K x UwSlowLen_Pls)    *)
(* K not learned / UwSlow_at_D_Req OFF -> fixed UwSlow_at_D_Val as before.  *)
(* Latched: once slowed down, the point is frozen (+10 mm hysteresis), so  *)
(* the lower speed does not move it back and speed up again. Released by   *)
(* a new roll (diameter 30 mm above the frozen point).                     *)

IF UwSlow_at_D_Req AND (RwMat_K > 0.0) AND (UwStopDiam_Limit > 0.0)
   AND (UwSlowLen_Pls > 0.0) THEN
    SqrtArg := UwStopDiam_Limit * UwStopDiam_Limit + 2.0 * RwMat_K * UwSlowLen_Pls;
    UwSlowDiamCalc := SQRT(SqrtArg);               (* same pattern as 6b *)
ELSE
    UwSlowDiamCalc := UwSlow_at_D_Val;
END_IF;

IF UwSlowDiamCalc < UwStopDiam_Limit + 10.0 THEN
    UwSlowDiamCalc := UwStopDiam_Limit + 10.0;
ELSIF UwSlowDiamCalc > 1500.0 THEN
    UwSlowDiamCalc := 1500.0;
END_IF;

IF UwSlowDiamLatch AND (UwDiam_Act > UwSlowDiamAct + 30.0) THEN
    UwSlowDiamLatch := FALSE;                       (* new roll *)
END_IF;

IF NOT UwSlowDiamLatch THEN
    UwSlowDiamAct := UwSlowDiamCalc;                (* live point, HMI *)
    IF Measure_ON AND (UwDiam_Act > 0.0) AND (UwDiam_Act <= UwSlowDiamCalc) THEN
        UwSlowDiamLatch := TRUE;
        UwSlowDiamAct := UwSlowDiamCalc + 10.0;     (* frozen + hysteresis *)
    END_IF;
END_IF;

(* ---- 7. Rewinder requests: latched, reset when a new core is loaded ---- *)

IF NOT RwStopEnable
   OR ((RwDiam < RwTargetDiam - RwResetHyst) AND NOT RwSensFault) THEN
    RwStop_at_D_Req := FALSE;
    RwSlow_at_D_Req := FALSE;
END_IF;

IF RwStopEnable THEN
    IF (RwRemain_Pls <= StopLen_Pls) OR (RwSensFault AND RwStopOnFault) THEN
        RwStop_at_D_Req := TRUE;
    END_IF;
    IF RwUseSlow AND (RwRemain_Pls <= RwSlowLen_Pls) THEN
        RwSlow_at_D_Req := TRUE;
    END_IF;
	
    (* v6t: thickness not learned (RwMat_K = 0): slow down at a fixed      *)
    (* distance before the target instead of stopping from full speed.    *)
	
    IF RwUseSlow AND (RwMat_K <= 0.0) AND (RwSlowFallbackMm > 0.0)
       AND NOT RwSensFault
       AND (RwDiam >= RwTargetDiam - RwSlowFallbackMm) THEN
        RwSlow_at_D_Req := TRUE;
    END_IF;
END_IF;

(* ---- 8. One AUTO at a time + single "SLOW DOWN AT" display ------------- *)

// ---- Refuse AUTO STOP when its target is already reached (HMI warning 20) ----
// AutoEnWhy (HMI bits): 1 = unwinder metres already reached, 2 = rewinder roll >= target

IF I_AutoStop_OS AND RwStopEnable AND NOT RwArmMem AND NOT RwSensFault
   AND (RwTargetDiam > REAL#0.0) AND (RwDiam >= RwTargetDiam - RwResetHyst) THEN
    RwStopEnable := FALSE;                          // refused
    AutoEnRefused := TRUE;
    AutoEnWhy := 2;
END_IF;

IF I_AutoStop_OS AND UwStopEnable AND NOT UwArmMem
   AND (UwStop_at_M_Val > REAL#0.0) AND (Current_Metre >= UwStop_at_M_Val) THEN
    UwStopEnable := FALSE;                          // refused
    AutoEnRefused := TRUE;
    AutoEnWhy := 1;
END_IF;

IF UwStopEnable AND NOT UwEnMem THEN                (* unwinder AUTO switched ON *)
    RwStopEnable := FALSE;
END_IF;

IF RwStopEnable AND NOT RwEnMem THEN                (* rewinder AUTO switched ON *)
    UwStopEnable := FALSE;
END_IF;

T_AutoEnRef(In := AutoEnRefused, PT := T#5s);       // warning shown 5 s

IF T_AutoEnRef.Q OR I_RsetAlarm OR Alarm_Reset THEN
    AutoEnRefused := FALSE;
END_IF;

RwArmMem := I_AutoStop_OS AND RwStopEnable;         // armed = selector 12SA5 AND enable
UwArmMem := I_AutoStop_OS AND UwStopEnable;
UwEnMem := UwStopEnable;
RwEnMem := RwStopEnable;

IF RwStopEnable THEN
    SlowAtDisp := RwSlow_at_D_Val;                     (* mm *)
    SlowAtMode := 2;
ELSIF UwStopEnable THEN
    SlowAtDisp := UwSlow_at_M_Val;                  (* m  *)
    SlowAtMode := 1;
ELSE
    SlowAtDisp := 0.0;
    SlowAtMode := 0;                                (* hide display *)
END_IF;

SlowAtShow := (SlowAtMode <> 0);

(* V11: unwinder column, same place, 3 states:                           *)
(*   AUTO STOP UNWINDER (12SA5 + unwinder AUTO) -> STOP LENGTH [m]       *)
(*   normal run, before the slow-down          -> SLOW AT Ø [mm]          *)
(*   slow-down reached (decel / final speed)   -> STOP AT Ø [mm]          *)
(* V11: stop by diameter EARLIER, so the web is stopped AT UwStopDiam_Limit:   *)
(* the stop command comes at UwStop_at_D_Val = UwStopDiam_Limit + the diameter   *)
(* of the paper unwound during the stop from the ACTUAL speed            *)
(* (StopLen_Pls, section 6, learned stop decel):                         *)
(*   UwStop_at_D_Val = SQRT(UwStopDiam_Limit^2 + 2 x RwMat_K x StopLen_Pls)       *)
(* General rung 18 (UwStopByDiam) compares with UwStop_at_D_Val.           *)
(* K not learned -> UwStopDiam_Limit (as before). Max UwStopDiam_Limit + 100 mm.     *)

UwStopLenShow  := I_AutoStop_OS AND UwStopEnable;
UwSlowDiamShow := NOT UwStopLenShow AND Measure_ON AND NOT UwSlowDiamLatch;
UwStopDiamShow := NOT UwStopLenShow AND Measure_ON AND UwSlowDiamLatch;

IF (RwMat_K > 0.0) AND (StopLen_Pls > 0.0) THEN
    SqrtArg := UwStopDiam_Limit * UwStopDiam_Limit + 2.0 * RwMat_K * StopLen_Pls;
    UwStop_at_D_Val := SQRT(SqrtArg);
ELSE
    UwStop_at_D_Val := UwStopDiam_Limit;
END_IF;

IF UwStop_at_D_Val > UwStopDiam_Limit + 100.0 THEN
    UwStop_at_D_Val := UwStopDiam_Limit + 100.0;
ELSIF UwStop_at_D_Val < UwStopDiam_Limit THEN
    UwStop_at_D_Val := UwStopDiam_Limit;
END_IF;

(* ---- 9. Automatic stop master = selector 12SA5 (I_AutoStop_OS) -------- *)

AutoSlowCmd := I_AutoStop_OS AND
               ((UwStopEnable AND UwSlow_at_M_Req) OR (RwStopEnable AND RwSlow_at_D_Req));

AutoStopCmd := I_AutoStop_OS AND
               ((UwStopEnable AND (UwStop_at_M_Val > 0.0)
                 AND (Current_Metre >= UwStop_at_M_Val))
                OR (RwStopEnable AND RwStop_at_D_Req));

(* ---- 10. Unwinder roll empty (for alarm 15) ---------------------------- *)

IF UwDiam_Act > (UwStopDiam_Limit + UwEmptyHyst) THEN
    UnWinder_Empty := FALSE;                        (* new roll loaded *)
END_IF;

IF (UwDiam_Act > 0.0) AND (UwDiam_Act <= UwStopDiam_Limit) THEN
    UnWinder_Empty := TRUE;                         (* roll empty *)
END_IF;

(* v6x: new parent roll loaded (empty -> not empty) -> HMI popup         *)

(* "DID YOU CHANGE THE PAPER (GSM)?". YES = forget the learned thickness *)
(* (same as NEW PAPER), NO = the HMI resets GsmAsk.                      *)
(* V9: ask only ONCE per REAL new roll: the roll must have been empty for *)
(* 3 s (arms the question), then the new roll must read more than        *)
(* UwStopDiam_Limit + 100 mm for 3 s. The sonar bouncing around UwStopDiam_Limit     *)
(* (empty core, hands, arms) no longer re-opens the popup.               *)

IF Tick THEN
    IF UnWinder_Empty THEN
		
        IF UwEmptyTicks < 1000 THEN
            UwEmptyTicks := UwEmptyTicks + 1;
        END_IF;
		
        IF UwEmptyTicks >= 30 THEN
            GsmArmed := TRUE;
        END_IF;
		
        UwFullTicks := 0;
    ELSE
        UwEmptyTicks := 0;
		
        IF GsmArmed AND Measure_ON AND (UwDiam_Act > UwStopDiam_Limit + 100.0) THEN
            UwFullTicks := UwFullTicks + 1;
			
            IF UwFullTicks >= 30 THEN
                GsmAsk := TRUE;
                GsmArmed := FALSE;
                UwFullTicks := 0;
            END_IF;
        ELSE
            UwFullTicks := 0;
        END_IF;
    END_IF;
END_IF;

UwEmptyMem := UnWinder_Empty;

IF GsmAskYes THEN
    RwMat_K := 0.0;
    RwMatLocked := FALSE;                           (* V9 *)
    LongActive := FALSE;
    LearnFailCnt := 0;
    MatChangeCnt := 0;
    GsmAskYes := FALSE;
    GsmAsk := FALSE;
END_IF;

(* V10: HMI popup "UNWINDER DIAMETER SENSOR SONAR IS OFF ! DO YOU WANT TO  *)
(* TURN IT ON ?" - only at standstill: at power-up and after every stop    *)
(* while Measure_ON = FALSE. YES (SonarAskYes, PLC resets it) = sonar ON;  *)
(* NO = the HMI resets SonarAsk (asked again after the next stop).         *)

IF Measure_ON THEN
    SonarAsk := FALSE;                              (* sonar ON: no popup *)
ELSIF NOT StartMotor_Cmd AND (SonarRunMem OR NOT SonarInit) THEN
    SonarAsk := TRUE;                               (* stopped / power-up *)
END_IF;

SonarInit := TRUE;
SonarRunMem := StartMotor_Cmd;

IF StartMotor_Cmd THEN
    SonarAsk := FALSE;                              (* never while running *)
END_IF;

IF SonarAskYes THEN
    Measure_ON := TRUE;
    SonarAsk := FALSE;
    SonarAskYes := FALSE;
END_IF;

(* ---- 11. Rewinder max diameter protection - ALWAYS active ------------- *)
(* Independent of selector 12SA5 and of the AUTO buttons.                  *)
(* Mechanical limit 680 mm radius = 1360 mm                                *)

IF NOT RwSensFault THEN
    RwLastValidDiam := RwDiam;
END_IF;

IF RwDiam >= RwMaxDiam THEN
    RwRemainMax_Pls := 0.0;
ELSIF RwMat_K > 0.0 THEN
    RwRemainMax_Pls := (RwMaxDiam * RwMaxDiam - RwDiam * RwDiam)
                       / (2.0 * RwMat_K);
ELSE
    RwRemainMax_Pls := 1.0E9;                       (* K not learned: plain limit *)
END_IF;

(* Display: diameter where the max-protection slow-down will start         *)

IF RwMat_K > 0.0 THEN
    SqrtArg := RwMaxDiam * RwMaxDiam - 2.0 * RwMat_K * RwSlowLen_Pls;
    IF SqrtArg > 0.0 THEN
        RwMaxSlowAtDiam := SQRT(SqrtArg);
    ELSE
        RwMaxSlowAtDiam := 0.0;
    END_IF;
ELSIF RwMaxSlowFallback > 0.0 THEN
    RwMaxSlowAtDiam := RwMaxSlowFallback;           (* fallback in use *)
ELSE
    RwMaxSlowAtDiam := RwMaxDiam;
END_IF;

(* Reset only after the roll is removed (diameter well below the limit)    *)

IF (RwDiam < RwMaxDiam - RwResetHyst) AND NOT RwSensFault THEN
    RwMaxStop := FALSE;
    RwMaxSlow := FALSE;
END_IF;

IF NOT RwSensFault THEN
	
    IF RwRemainMax_Pls <= StopLen_Pls THEN
        RwMaxStop := TRUE;                          (* speed-compensated stop *)
    END_IF;
	
    IF RwRemainMax_Pls <= RwSlowLen_Pls THEN
        RwMaxSlow := TRUE;                          (* warning slow-down + horn *)
    END_IF;
	
    IF (RwMat_K <= 0.0) AND (RwMaxSlowFallback > 0.0)
       AND (RwDiam >= RwMaxSlowFallback) THEN
        RwMaxSlow := TRUE;                          (* fallback while K not learned *)
    END_IF;
	
ELSIF (AI_Diam_Rewinder < RwRawMin) AND (RwLastValidDiam > RwMaxDiam - 100.0) THEN
    RwMaxStop := TRUE;                              (* roll grew into the DT35 near zone *)
END_IF;

(* Max diameter protection added OUTSIDE the 12SA5 master (section 9)      *)

AutoSlowCmd := AutoSlowCmd OR RwMaxSlow;
AutoStopCmd := AutoStopCmd OR RwMaxStop;

(* ---- 11b. V12: END-OF-ROLL STOP RAMP ---------------------------------- *)
(* Normal end-of-roll stops (AutoStopCmd: unwinder metres, rewinder target,*)
(* rewinder max diameter; UwStopByDiam: unwinder diameter) no longer drop  *)
(* the run command at once (drive DEC ramp 3 s = 20 Hz/s -> up to 8 m/s2  *)
(* of web on a big roll, hard on the rewinder gearbox). With the feed-    *)
(* forward in AUTO they start the SOFT STOP at FinalStopDecel (General    *)
(* rung 10); the run command drops below SoftStopEndSpd. START cannot     *)
(* cancel it. The stop lengths (section 6) use the same ramp, so the web  *)
(* still stops at the target / UwStopDiam_Limit.                          *)
(* Immediate stop (EndStopNow -> Motor_Manager rung 4 Stop):              *)
(*   ramp not usable (FinalStopDecel 0, FFEnable OFF, ManMode, JOG, the    *)
(*   motor stopped = start blocked as before), or safety net: unwinder    *)
(*   10 mm below UwStopDiam_Limit / rewinder at RwMaxDiam during the ramp.*)

IF FinalStopDecel < 0.0 THEN
    FinalStopDecel := 0.0;
ELSIF (FinalStopDecel > 0.0) AND (FinalStopDecel < 50.0) THEN
    FinalStopDecel := 50.0;
ELSIF FinalStopDecel > 2000.0 THEN
    FinalStopDecel := 2000.0;
END_IF;

EndStopReq := AutoStopCmd OR (Measure_ON AND UwStopByDiam);
EndRampOK := (FinalStopDecel > 0.0) AND FFActive AND StartMotor_Cmd;

IF EndStopReq AND EndRampOK THEN
    FinalStopRamp := TRUE;                          (* -> soft stop, General 10 *)
END_IF;

IF NOT StartMotor_Cmd THEN
    FinalStopRamp := FALSE;
END_IF;

EndRampHard := FinalStopRamp
               AND ((Measure_ON AND (UwDiam_Act > 0.0)
                     AND (UwDiam_Act < UwStopDiam_Limit - 10.0))
                    OR ((RwDiam >= RwMaxDiam) AND NOT RwSensFault));

EndStopNow := (EndStopReq AND NOT FinalStopRamp) OR EndRampHard;

// ---- 11c. Auto stop DONE (HMI warning 19), latched until START / RESET ----
// AutoStopWhy: 1 unwinder metres, 2 rewinder diameter, 4 rewinder MAX, 8 unwinder diameter

IF StartMotor_Cmd AND NOT AS_RunMem THEN           // new START: clear
    AutoStopDone := FALSE;
    AutoStopSeen := FALSE;
    AutoStopWhy := 0;
END_IF;

IF StartMotor_Cmd AND EndStopReq AND NOT AutoStopSeen THEN
    AutoStopSeen := TRUE;                           // auto stop started while running
	
    IF RwMaxStop THEN
        AutoStopWhy := 4;                           // rewinder MAX (protection, highest)
    ELSIF I_AutoStop_OS AND RwStopEnable AND RwStop_at_D_Req THEN
        AutoStopWhy := 2;                           // rewinder diameter reached
    ELSIF Measure_ON AND UwStopByDiam THEN
        AutoStopWhy := 8;                           // unwinder diameter (sonar)
    ELSE
        AutoStopWhy := 1;                           // unwinder metres
    END_IF;
END_IF;

IF AS_RunMem AND NOT StartMotor_Cmd AND AutoStopSeen THEN
    AutoStopDone := TRUE;                           // stopped by the auto stop
END_IF;

IF I_RsetAlarm OR Alarm_Reset THEN
    AutoStopDone := FALSE;
END_IF;

T_AutoStopDisp(In := AutoStopDone, PT := T#8s);    // show the warning 8s 

IF T_AutoStopDisp.Q THEN
    AutoStopDone := FALSE;
END_IF;

AS_RunMem := StartMotor_Cmd;

(* ---- 12. Learning supervision -> alarm 16 (section Alarms) ------------ *)
(* Learned paper thickness, for display / plausibility check               *)

IF MmPerPulse > 0.0 THEN
    RwThick_mm := RwMat_K * 3.14159 / (2.0 * MmPerPulse);
ELSE
    RwThick_mm := 0.0;
END_IF;

(* Fault: too many consecutive windows / stops that should have            *)
(* learned but did not. Clears by itself on the next good result.          *)
(* v6w: ALARM RESET (panel button or HMI) also clears the fail counters, *)
(* so alarm 16 resets in one press. It comes back only if the learning  *)
(* fails again RwLearnFailMax / RwStopFailMax times in a row.           *)

IF I_RsetAlarm OR Alarm_Reset THEN
    LearnFailCnt := 0;
    StopFailCnt := 0;
END_IF;

GSM_LearnFault := (LearnFailCnt >= RwLearnFailMax)
              OR (StopFailCnt >= RwStopFailMax);       (* -> alarm 16 *)

(* v6e: learning status for the HMI. FALSE until learned.                   *)

GSM_Learned_OK := (RwMat_K > 0.0)
                AND ((RwStopDecel > 0.0) OR NOT RwLearnStop)
                AND NOT GSM_LearnFault;

(* ---- 13. v6h: keep T-one in automatic tension control during the stop - *)
(* While running: BrakeHold = Brake_Cmd (no change in running behaviour).  *)
(* After the stop: stays ON until the web is below 5 m/min, after 15 s,   *)
(* or on E-stop. Already TRUE on the stop scan (Output_Manager runs before *)
(* this section), so O_Brake never drops for one scan.                     *)
(* Output_Manager rung 2:  O_Brake := Brake_Cmd OR BrakeHold               *)

IF O_MotorStart THEN
    BrakeHold := Brake_Cmd AND ControlVoltage;
    BrakeHoldTicks := 0;
ELSIF BrakeHold THEN
	
    IF Tick THEN
        BrakeHoldTicks := BrakeHoldTicks + 1;
    END_IF;
	
    (* v6v: signed web speed: a web pulled BACK (negative speed) also     *)
    (* releases the T-one (trace 10/28 15:00: -6.6 m/min, about 20 cm).  *)
	
    IF NOT ControlVoltage OR (Velocity_M_min < 5.0) OR (BrakeHoldTicks >= 150) THEN
        BrakeHold := FALSE;
    END_IF;
END_IF;

(* ---- 14. v6j: TEACH CORE - automatic offset with an empty core -------- *)
(* HMI: set RwTeachCore (button, Set ON). Conditions: motor stopped, web  *)
(* not moving, DT35 OK. After 2 s stable (filter settled):                 *)
(*     RwAxisDist := RwDist + RwCoreDiameter / 2   -> RwDiam = RwCoreDiameter          *)
(* RwTeachState: 0 idle, 1 teaching (wait 2 s), 2 done OK,                *)
(*               3 refused (motor running / web moving / DT35 fault).     *)
(* Only the offset is taught: the scale is RwDist10V - RwDist0V           *)
(* (= real distance between the two DT35 taught points).                  *)

IF RwTeachCore THEN
    IF O_MotorStart OR (RwSpeed > 1.0) OR RwSensFault
       OR NOT RwFiltInit OR (RwCoreDiameter <= 0.0) THEN
        RwTeachState := 3;                          (* refused *)
        RwTeachCore := FALSE;
        TeachTicks := 0;
    ELSE
        RwTeachState := 1;                          (* teaching *)
		
        IF Tick THEN
            TeachTicks := TeachTicks + 1;
        END_IF;
		
        IF TeachTicks >= 20 THEN                    (* 2 s stable *)
            RwAxisDist_Prev := RwAxisDist;          (* v6l: keep previous *)
            RwAxisDist := RwDist + RwCoreDiameter / 2.0;
            RwTeachState := 2;                      (* done *)
            RwTeachCore := FALSE;
            TeachTicks := 0;
        END_IF;
    END_IF;
ELSE
    TeachTicks := 0;
	
    IF O_MotorStart THEN
        RwTeachState := 0;                          (* clear status on next run *)
    END_IF;
END_IF;

(* ---- 14b. v6k: unwinder TEACH CORE (HMI button Core_Measure) ---------- *)
(* Same behaviour as section 14. Sonar is not filtered, so the 2 s are   *)
(* averaged:  UwCoreDistance := average(UwDiam_Measure)  (sonar -> core   *)
(* surface). UwDiam_Act = (UwCoreDistance - UwDiam_Measure) * 2           *)
(*                        + UwCoreDiameter   (General rung 14, unchanged). *)
(* UwTeachState: 0 idle, 1 teaching, 2 done OK, 3 refused.                 *)

IF Core_Measure THEN
	
    IF O_MotorStart OR (RwSpeed > 1.0) OR (UwCoreDiameter <= 0.0)
       OR (UwDiam_Measure <= 0.0) THEN
        UwTeachState := 3;                          (* refused *)
        Core_Measure := FALSE;
        UwTeachTicks := 0;
        UwTeachSum := 0.0;
    ELSE
        UwTeachState := 1;                          (* teaching *)
		
        IF Tick THEN
            UwTeachTicks := UwTeachTicks + 1;
            UwTeachSum := UwTeachSum + UwDiam_Measure;
        END_IF;
		
        IF UwTeachTicks >= 20 THEN                  (* 2 s, 20 samples *)
            UwCoreDist_Prev := UwCoreDistance;      (* v6l: keep previous *)
            UwCoreDistance := UwTeachSum / INT_TO_REAL(UwTeachTicks);
            UwTeachState := 2;                      (* done *)
            Core_Measure := FALSE;
            UwTeachTicks := 0;
            UwTeachSum := 0.0;
        END_IF;
    END_IF;
ELSE
    UwTeachTicks := 0;
    UwTeachSum := 0.0;
	
    IF O_MotorStart THEN
        UwTeachState := 0;                          (* clear status on next run *)
    END_IF;
END_IF;

(* ---- 14c. v6l: UNDO teach = swap current <-> previous (machine stopped) *)
(* Pressing UNDO twice goes back to the taught value. State 4 = RESTORED. *)

IF RwTeachUndo THEN
	
    IF NOT O_MotorStart AND (RwAxisDist_Prev > 0.0) THEN
        TeachSwap := RwAxisDist;
        RwAxisDist := RwAxisDist_Prev;
        RwAxisDist_Prev := TeachSwap;
        RwTeachState := 4;                          (* restored *)
    ELSE
        RwTeachState := 3;                          (* refused *)
    END_IF;
    RwTeachUndo := FALSE;
END_IF;

IF UwTeachUndo THEN
	
    IF NOT O_MotorStart AND (UwCoreDist_Prev > 0.0) THEN
        TeachSwap := UwCoreDistance;
        UwCoreDistance := UwCoreDist_Prev;
        UwCoreDist_Prev := TeachSwap;
        UwTeachState := 4;                          (* restored *)
    ELSE
        UwTeachState := 3;                          (* refused *)
    END_IF;
    UwTeachUndo := FALSE;
END_IF;

(* Section Tension_Helper: ladder, written here as Structured Text *)

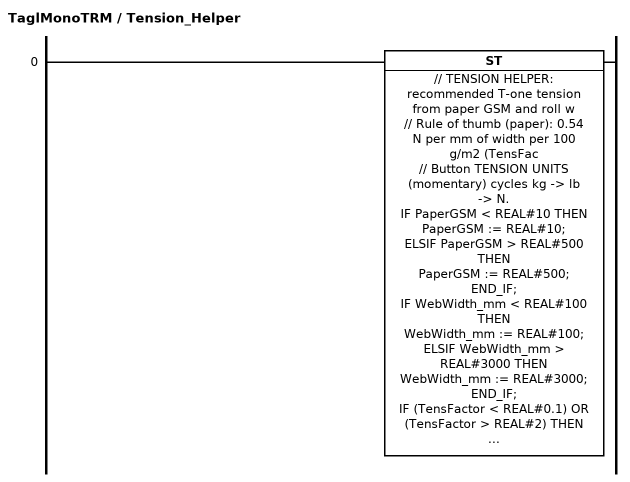
(* Rung 0 *)
// TENSION HELPER: recommended T-one tension from paper GSM and roll width.
// Rule of thumb (paper): 0.54 N per mm of width per 100 g/m2 (TensFactor).
// Button TENSION UNITS (momentary) cycles kg -> lb -> N.

IF PaperGSM < REAL#10 THEN
    PaperGSM := REAL#10;
ELSIF PaperGSM > REAL#500 THEN
    PaperGSM := REAL#500;
END_IF;

IF WebWidth_mm < REAL#100 THEN
    WebWidth_mm := REAL#100;
ELSIF WebWidth_mm > REAL#3000 THEN
    WebWidth_mm := REAL#3000;
END_IF;

IF (TensFactor < REAL#0.1) OR (TensFactor > REAL#2) THEN
    TensFactor := REAL#0.54;
END_IF;

// Unit button: one press = next unit

IF TensUnitPB AND NOT TensUnitMem THEN
    TensUnit := TensUnit + 1;
    IF TensUnit > 2 THEN
        TensUnit := 0;
    END_IF;
END_IF;

TensUnitMem := TensUnitPB;

IF (TensUnit < 0) OR (TensUnit > 2) THEN
    TensUnit := 0;
END_IF;

TensIdeal_N := PaperGSM / REAL#100 * WebWidth_mm * TensFactor;

CASE TensUnit OF
    1:  TensIdeal_Disp := TensIdeal_N / REAL#9.81 * REAL#2.20462;   // lb
    2:  TensIdeal_Disp := TensIdeal_N;                               // N
ELSE
        TensIdeal_Disp := TensIdeal_N / REAL#9.81;                   // kg
END_CASE;

TensShowKg := (TensUnit = 0);
TensShowLb := (TensUnit = 1);
TensShowN  := (TensUnit = 2);
END_PROGRAM